Fanuc KAREL source: ka00145.KL

-- PROVISIONAL review KL for V1013-1; original PC SHA256 22c2bfee81efff36ba0acade6bb1509a8c545dd202ea1ea47fc56999cd50d5f3
-- Incomplete behavior may be omitted. Consult companion uncertainty JSON. Do not deploy.
PROGRAM KA00145
%NOLOCKGROUP
-- UNRESOLVED_DECL SRC type=002010
-- UNRESOLVED_DECL DST type=002010
BEGIN
  -- UNRESOLVED_PC offsets 5-19; opcodes 22,22,1E
  -- UNRESOLVED_PC offsets 24-28; opcodes 7F
END KA00145
